Fanuc KAREL source: kt00891.KL

-- PROVISIONAL review KL for V1013-1; original PC SHA256 cafad1b3a2084525d2c0fc9fbf7a7c3586466ef35f94dd3eb4cb1401c935bbaa
-- Incomplete behavior may be omitted. Consult companion uncertainty JSON. Do not deploy.
PROGRAM KT00891
%NOLOCKGROUP
-- UNRESOLVED_DECL P1 type=000199
-- UNRESOLVED_DECL P2 type=000199
-- UNRESOLVED_DECL OUT type=000101
BEGIN
  -- UNRESOLVED_PC offsets 5-35; opcodes 27,27,49,7E,AD,76,7E,4A
  -- UNRESOLVED_PC offsets 40-44; opcodes 7F
END KT00891
